Fanuc KAREL source: ks00003.KL

-- PROVISIONAL review KL for V1013-1; original PC SHA256 5a57a0293546b7cc65f30ac3457deee017ab55689b94299437d7172972988f47
-- Incomplete behavior may be omitted. Consult companion uncertainty JSON. Do not deploy.
PROGRAM KS00003
%NOLOCKGROUP
VAR
  FLAG : BOOLEAN
  N : INTEGER
  STATUS : INTEGER
  PN : STRING[80]
  VN : STRING[80]
-- UNRESOLVED_DECL A type=001100
-- UNRESOLVED_DECL B type=001100
BEGIN
  -- UNRESOLVED_PC offsets 5-13; opcodes 3F,75
  -- UNRESOLVED_PC offsets 18-27; opcodes 3F,75
  -- UNRESOLVED_PC offsets 32-47; opcodes 22,22,30
  -- UNRESOLVED_PC offsets 52-56; opcodes 7F
END KS00003
